Fanuc KAREL source: KT00687.KL

PROGRAM KT00687
%NOLOCKGROUP
VAR
  P1: JOINTPOS
  P2: JOINTPOS
  OUT: BOOLEAN
BEGIN
  OUT = - P1
END KT00687
